(* IEC 61131-3 sources: Lasal-MCP/examples/SampleSource/LASALScreenAdvancedSolution/LASALScreenAdvancedSolution/LASALScreenAdvacnedSolution/Stations/Terminal/HMI/Network/ExamplesNet, 1 file *)

(* ---- ONE_ExamplesNet_Table.st ---- *)
#define OBJECTS_CONFIG

#include <.\lsl_st_mt.h>

FUNCTION GLOBAL TAB ONE_ExamplesNet
-1$UINT, 0$UINT,
0$UINT, 0$UINT,

11$UDINT,
TO_UDINT(2980745877), "_MyIO", 0$UINT, 3$UINT, 0$UINT,
TO_UDINT(1412211373), "DataRecord", 0$UINT, 0$UINT, 1$UINT,
TO_UDINT(1396269567), "DataRecordSave", 0$UINT, 0$UINT, 1$UINT,
TO_UDINT(2984478465), "FileHandling", 0$UINT, 0$UINT, 1$UINT,
TO_UDINT(1011632712), "FileRead", 0$UINT, 0$UINT, 1$UINT,
TO_UDINT(2515960668), "Indicator", 0$UINT, 0$UINT, 1$UINT,
TO_UDINT(2225119864), "MerkerEx", 1$UINT, 22$UINT, 0$UINT,
TO_UDINT(933570811), "RAMex", 1$UINT, 17$UINT, 4$UINT,
TO_UDINT(2898603620), "StringInternal", 1$UINT, 84$UINT, 0$UINT,
TO_UDINT(2408581120), "StringRAM", 1$UINT, 10$UINT, 4$UINT,
TO_UDINT(3232495061), "VirtualBaseInit", 1$UINT, 3$UINT, 0$UINT,

_NO_ATTR, TO_UDINT(737090624), "DATARECORD1",

_NO_ATTR, TO_UDINT(2928490843), "DATARECORDSAVE1",

_NO_ATTR, TO_UDINT(4100603046), "FILEHANDLING1",

_NO_ATTR, TO_UDINT(4226247263), "FILEREAD1",

_NO_ATTR, TO_UDINT(3784574187), "INDICATOR1",

1$UINT, TO_UDINT(2770400313), "FILEHANDLING1\DRIVENAME\DATABUFFER",
1$UINT, TO_UDINT(4027332554), "FILEHANDLING1\FILEEXTENSION\DATABUFFER",
1$UINT, TO_UDINT(3113375051), "FILEHANDLING1\FILENAME\DATABUFFER",
1$UINT, TO_UDINT(1504833645), "STRINGRAM1\DATABUFFER",

1$UINT, TO_UDINT(3139633982), "FILEHANDLING1\DRIVENAME",
1$UINT, TO_UDINT(624134213), "FILEHANDLING1\FILEEXTENSION",
1$UINT, TO_UDINT(158136700), "FILEHANDLING1\FILENAME",
_NO_ATTR, TO_UDINT(2203287487), "STRINGRAM1",

//Internal connections
0$UDINT,
7$UDINT,
TO_UDINT(2), "DriveName", TO_UDINT(9),
TO_UDINT(2), "FileName", TO_UDINT(11),
TO_UDINT(2), "FileExtension", TO_UDINT(10),
TO_UDINT(9), "DataBuffer", TO_UDINT(5),
TO_UDINT(10), "DataBuffer", TO_UDINT(6),
TO_UDINT(11), "DataBuffer", TO_UDINT(7),
TO_UDINT(12), "DataBuffer", TO_UDINT(8),
0$UDINT,
8$UDINT,
TO_UDINT(1), "FileRead", TO_UDINT(3), "ReadSteps",
TO_UDINT(1), "FileHandling", TO_UDINT(2), "Steps",
TO_UDINT(2), "FileRead", TO_UDINT(3), "ReadSteps",
TO_UDINT(3), "StringRAM", TO_UDINT(12), "Data",
TO_UDINT(9), "DataBuffer", TO_UDINT(5), "m_udLength",
TO_UDINT(10), "DataBuffer", TO_UDINT(6), "m_udLength",
TO_UDINT(11), "DataBuffer", TO_UDINT(7), "m_udLength",
TO_UDINT(12), "DataBuffer", TO_UDINT(8), "m_udLength",

//Initialization values
0$UDINT,
10$UDINT,
TO_UDINT(0), "AllocateSize", TO_UDINT(4 KB),//|ExamplesNet.DataRecord1.AllocateSize;
TO_UDINT(1), "AllocateSize", TO_UDINT(4 KB),//|ExamplesNet.DataRecordSave1.AllocateSize;
TO_UDINT(5), "ThreadSafe", TO_UDINT(0),//|ExamplesNet.DriveName\FileHandling1\DataBuffer.ThreadSafe;
TO_UDINT(6), "ThreadSafe", TO_UDINT(0),//|ExamplesNet.FileExtension\FileHandling1\DataBuffer.ThreadSafe;
TO_UDINT(7), "ThreadSafe", TO_UDINT(0),//|ExamplesNet.FileName\FileHandling1\DataBuffer.ThreadSafe;
TO_UDINT(8), "ThreadSafe", TO_UDINT(0),//|ExamplesNet.StringRAM1\DataBuffer.ThreadSafe;
TO_UDINT(9), "SingleRealloc", TO_UDINT(1),//|ExamplesNet.FileHandling1\DriveName.SingleRealloc;
TO_UDINT(10), "SingleRealloc", TO_UDINT(1),//|ExamplesNet.FileHandling1\FileExtension.SingleRealloc;
TO_UDINT(11), "SingleRealloc", TO_UDINT(1),//|ExamplesNet.FileHandling1\FileName.SingleRealloc;
TO_UDINT(12), "SingleRealloc", TO_UDINT(1),//|ExamplesNet.StringRAM1.SingleRealloc;

//Symbolic initialization values
0$UDINT,
0$UDINT,

//Initialization of string values
0$UDINT,
4$UDINT,
TO_UDINT(9), "", 0$UINT, TO_UINT(OFF(L1)-OFF(L0)), L0:"C:\",L1://|ExamplesNet.FileHandling1\DriveName.Data;
TO_UDINT(10), "", 0$UINT, TO_UINT(OFF(L3)-OFF(L2)), L2:".txt",L3://|ExamplesNet.FileHandling1\FileExtension.Data;
TO_UDINT(11), "", 0$UINT, TO_UINT(OFF(L5)-OFF(L4)), L4:"MyFile",L5://|ExamplesNet.FileHandling1\FileName.Data;
TO_UDINT(12), "", 0$UINT, TO_UINT(OFF(L7)-OFF(L6)), L6:"C:\MyFile.txt",L7://|ExamplesNet.StringRAM1.Data;

//Configuration of tasks (RealTime, Cyclic, Background)
0$UDINT,
0$UDINT,

0$UDINT,
0$UDINT,

0$UDINT,
2$UDINT,
TO_UDINT(2), (50)$UDINT, 4194303$DINT, 	//FILEHANDLING1
TO_UDINT(3), (10)$UDINT, 4194303$DINT, 	//FILEREAD1

//External connections
0$UDINT,
3$UDINT,
TO_UDINT(0), "Lse", C_DIR, TO_UDINT(299963966), "Lse","Lse",
TO_UDINT(1), "Lse", C_DIR, TO_UDINT(299963966), "Lse","Lse",
TO_UDINT(4), "Lse", C_DIR, TO_UDINT(299963966), "Lse","Lse",

//Magic internal connections
0$UDINT,
4$UDINT,
TO_UDINT(5), "UseFile", TO_UDINT(9), "UseFile",
TO_UDINT(6), "UseFile", TO_UDINT(10), "UseFile",
TO_UDINT(7), "UseFile", TO_UDINT(11), "UseFile",
TO_UDINT(8), "UseFile", TO_UDINT(12), "UseFile",

//Configuration of timeslots of tasks (RealTime, Cyclic)
#ifdef __LSLLDR_TIMESLOTS__
0$UDINT,
0$UDINT,

0$UDINT,
0$UDINT,

#endif //__LSLLDR_TIMESLOTS__

//MultiMaster connections
#ifdef __LSLLDR_MULTIMASTER__
0$UDINT,
0$UDINT,
#endif //__LSLLDR_MULTIMASTER__

//Configuration for task ID (RealTime, CyclicTime)
#ifdef __LSLLDR_TASKID__
"\\\\TASKS2  "
0$UDINT,
0$UDINT,

0$UDINT,
0$UDINT,

0$UDINT,
2$UDINT,
(0)$UDINT, 	//FILEHANDLING1
(0)$UDINT, 	//FILEREAD1

#endif //__LSLLDR_TASKID__

END_FUNCTION
